Fanuc KAREL source: KT00144.KL

PROGRAM KT00144
%NOLOCKGROUP
VAR
  R1: REAL
  H2: ARRAY[2] OF SHORT
  OUT: REAL
BEGIN
  R1 = 2.0
    H2[1] = 3
  OUT = R1 DIV H2[1]
END KT00144
